RoboDK station: paint_booth.rdk

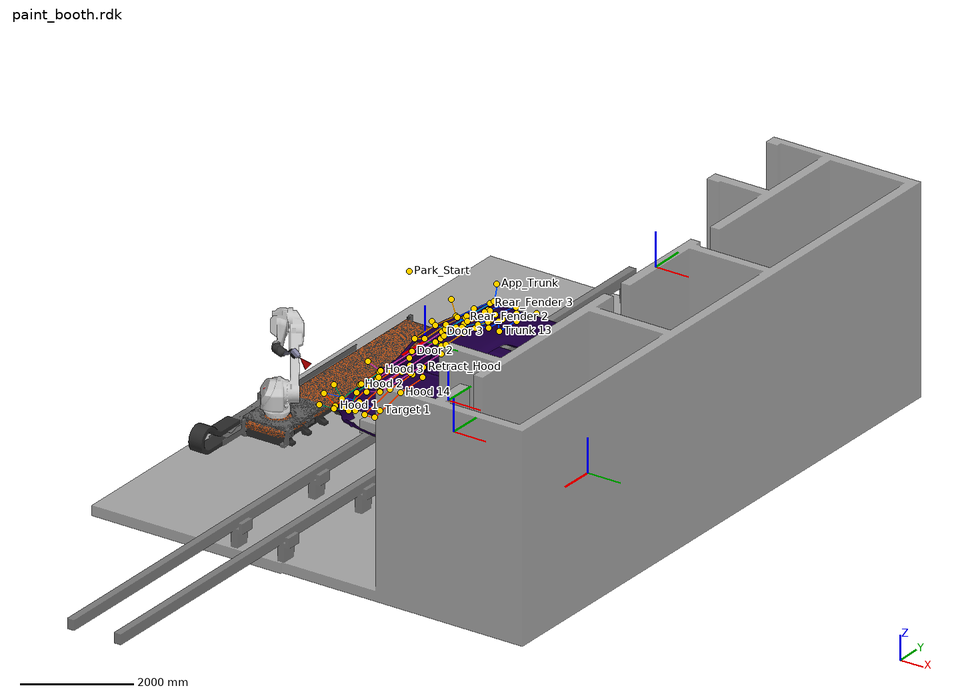
[picture v0: the station drawn from its stored meshes, robots at their saved joint values, targets as dots, program paths as lines]
Station paint booth backup2 (saved by RoboDK 6.1.1). Poses are relative to the parent item; angles as X-Y-Z fixed-axis rotations.
Station parameters (name, value as stored): AttachCamera_Record, 1, Record_Record, 0
  - frame ABB IRBT 7004 Standard 4m Base at (0, 2700, 0) mm, rotated rx 0 ry 0 rz -90 deg
    - robot ABB IRBT 7004 Standard 4m: 1 axes
        modified DH rows (alpha deg, a mm, theta deg, d mm): 0, 0, 0, 0 linear
        base shift (840.5, 4.2, 379.5) mm, rotated rx 0 ry 90 rz 0 deg
        joint limits [0] to [3700]; home [0]; saved at [3700]
      - robot ABB IRB 5500-27: 6 axes, payload 16 kg, reach 2200 mm, repeatability 0.15 mm, weight 600 kg
          modified DH rows (alpha deg, a mm, theta deg, d mm): 0, 0, 0, 436; -90, 0, -90, -5; 0, 1300, 0, 0; -90, 0, -90, 1510.5; 35, 0, 0, 79.169; -70, 0, 180, 79.169
          base shift (0, 0, 0) mm, rotated rx 0 ry 0 rz 90 deg
          joint limits [-104, -65, -70, -719, -719, -720] to [104, 150, 70, 719, 719, 720]; home [0, 0, 0, 0, 0, 0]; saved at [-54.839, -32.896, 27.054, 12.85, -64.516, 53.554]
        - tool Generic Paint Sprayer, TCP at (87.9, 0, 515.6) mm, rotated rx 0 ry 30 rz 0 deg, size 277.6 x 203.2 x 501.7 mm
  - frame booth_frame at (5380, 0, 0) mm, rotated rx 0 ry 0 rz -90 deg
    - folder Paint_Booth
      - object paint booth v1_paint booth v1_Back wall at (0, 0, 0) mm, size 12200 x 2000 x 4000 mm, geometry from paint booth v1_paint booth v1_Back wall.stl
      - object paint booth v1_paint booth v1_entry_part at (0, 0, 0) mm, size 250 x 1150 x 4000 mm, geometry from paint booth v1_paint booth v1_entry_part.stl
      - object paint booth v1_paint booth v1_entry_wall (1) at (0, 0, 0) mm, size 250 x 1150 x 4000 mm, geometry from paint booth v1_paint booth v1_entry_wall (1).stl
      - object paint booth v1_paint booth v1_entry_wall at (0, 0, 0) mm, size 1700 x 439.1 x 4000 mm, geometry from paint booth v1_paint booth v1_entry_wall.stl
      - object paint booth v1_paint booth v1_exit_wall (1) at (0, 0, 0) mm, size 250 x 1150 x 4000 mm, geometry from paint booth v1_paint booth v1_exit_wall (1).stl
      - object paint booth v1_paint booth v1_exit_wall (2) at (0, 0, 0) mm, size 250 x 1150 x 4000 mm, geometry from paint booth v1_paint booth v1_exit_wall (2).stl
      - object paint booth v1_paint booth v1_exit_wall at (0, 0, 0) mm, size 2500 x 439.1 x 4000 mm, geometry from paint booth v1_paint booth v1_exit_wall.stl
      - object paint booth v1_paint booth v1_floor at (0, 0, 0) mm, size 12240.8 x 9200 x 200 mm, geometry from paint booth v1_paint booth v1_floor.stl
      - object paint booth v1_paint booth v1_front_wall at (0, 0, 0) mm, size 8000 x 200 x 4000 mm, geometry from paint booth v1_paint booth v1_front_wall.stl
      - object paint booth v1_paint booth v1_mid_wall (1) at (0, 0, 0) mm, size 4000 x 200 x 4000 mm, geometry from paint booth v1_paint booth v1_mid_wall (1).stl
      - object paint booth v1_paint booth v1_mid_wall (2) at (0, 0, 0) mm, size 950 x 200 x 4000 mm, geometry from paint booth v1_paint booth v1_mid_wall (2).stl
      - object paint booth v1_paint booth v1_mid_wall (3) at (0, 0, 0) mm, size 3400 x 200 x 4000 mm, geometry from paint booth v1_paint booth v1_mid_wall (3).stl
      - object paint booth v1_paint booth v1_mid_wall at (0, 0, 0) mm, size 2150 x 200 x 4000 mm, geometry from paint booth v1_paint booth v1_mid_wall.stl
  - frame conveyor_frame at (2500, 0, 0) mm
    - object Conveyor at (0, 6191.19, 0) mm, rotated rx 0 ry 0 rz -90 deg, size 17200 x 1350 x 600 mm, geometry from Conveyor.stl
    - object cart at (0, 6191.19, 0) mm, size 1500 x 3500 x 250 mm, geometry from cart.stl
    - frame frame_base at (0, 6191.19, 750) mm
    - target Conv_Entry (joint target) at (0, 1691.19, 750) mm; joints [0] of Conveyor
    - target Conv_Paint (joint target) at (0, 1691.19, 750) mm; joints [4500] of Conveyor
    - target Conv_Exit (joint target) at (0, 1691.19, 750) mm; joints [13248.192] of Conveyor
  - frame Conveyor at (2500, 6191.19, 750) mm
    - robot Conveyor: 1 axes
        modified DH rows (alpha deg, a mm, theta deg, d mm): 0, 0, 0, 0 linear
        base shift (0, 0, 0) mm, rotated rx 90 ry 0 rz 0 deg
        joint limits [0] to [15000]; home [0]; saved at [4500]
      - frame car_frame at (0, -1850, -70) mm
        - object car_body at (0, 0, 0) mm, rotated rx 90 ry 0 rz 90 deg, size 4801.1 x 1114.9 x 1961.6 mm, geometry from car_body_optimised.obj
        - target Target 1 (Cartesian target) at (20.58, -2128.6, 648.13) mm, rotated rx 159.32 ry 5.46 rz -156.1 deg; joints [-17.994, 40.195, -43.091, -41.526, -55.736, 93.269, 3700] of ABB IRB 5500-27
        - target Target 2 (Cartesian target) at (-499.07, -2013.93, 637.53) mm, rotated rx 169.55 ry 9.47 rz -156.84 deg; joints [-17.854, 10.002, -1.972, -48.865, -37.872, 74.599, 3700] of ABB IRB 5500-27
        - object car_paint_1 at (-2500, 158.81, -680) mm, size 1941.7 x 1314.7 x 689.4 mm
        - object car_paint_2 at (-2500, 158.81, -680) mm, size 1932.4 x 3061.3 x 1113.1 mm
        - object car_paint_3 at (-2500, 158.81, -680) mm, size 1960.3 x 2051 x 1094.9 mm
        - object car_paint_4 at (-2500, 158.81, -680) mm, size 1961.6 x 1256.6 x 838.3 mm
        - target Hood 1 (Cartesian target) at (-850, -2240, 549.52) mm, rotated rx 170.58 ry 46.52 rz 180 deg; joints [-33.908, -9.39, 33.602, 38.78, -64.314, 10.994, 3700] of ABB IRB 5500-27
        - target Hood 2 (Cartesian target) at (-850, -1495, 668.46) mm, rotated rx 175.62 ry 0.84 rz -135.11 deg; joints [-8.251, -3.639, 8.764, -39.401, -59.237, 68.878, 3513] of ABB IRB 5500-27
        - target Hood 3 (Cartesian target) at (-850, -850, 690.55) mm, rotated rx 179.29 ry 0.3 rz -135 deg; joints [-7.072, -4.967, 9.136, -44.55, -55.783, 68.456, 2868] of ABB IRB 5500-27
        - target Hood 4 (Cartesian target) at (-625, -850, 729.52) mm, rotated rx -176.51 ry 5.77 rz -134.73 deg; joints [-6.745, 1.906, 2.143, -43.43, -50.492, 62.325, 2868] of ABB IRB 5500-27
        - target Hood 5 (Cartesian target) at (-625, -1505, 702.48) mm, rotated rx 179.51 ry 6.71 rz -134.83 deg; joints [-8.01, 3.25, 1.791, -36.982, -54.709, 62.353, 3523] of ABB IRB 5500-27
        - target Hood 6 (Cartesian target) at (-625, -2260, 584.84) mm, rotated rx 153.99 ry 5.37 rz -180 deg; joints [-27.175, 8.933, 2.732, -74.826, -17.731, 103.498, 3700] of ABB IRB 5500-27
        - target Hood 7 (Cartesian target) at (-400, -2280, 595.96) mm, rotated rx 166.53 ry -24.84 rz 109.32 deg; joints [-16.554, 21.687, -16.957, -133.314, -63.434, 218.22, 3700] of ABB IRB 5500-27
        - target Hood 8 (Cartesian target) at (-400, -1515, 725.47) mm, rotated rx 177.2 ry 3.28 rz 134.91 deg; joints [6.733, 12.58, -7.202, -178.41, -50.579, 227.726, 3533] of ABB IRB 5500-27
        - target Hood 9 (Cartesian target) at (-400, -850, 782.15) mm, rotated rx 177.63 ry 2.98 rz 134.92 deg; joints [6.843, 12.694, -9.476, -174.35, -52.852, 224.109, 2868] of ABB IRB 5500-27
        - target Hood 10 (Cartesian target) at (-175, -850, 793.95) mm, rotated rx 179.19 ry 2.16 rz 134.97 deg; joints [6.345, 23.93, -24.263, -167.605, -56.502, 217.205, 2868] of ABB IRB 5500-27
        - target Hood 11 (Cartesian target) at (-175, -1535, 771.67) mm, rotated rx 175.02 ry -3.19 rz 135.2 deg; joints [4.513, 24.031, -24.527, -162.354, -53.815, 216.084, 3553] of ABB IRB 5500-27
        - target Hood 12 (Cartesian target) at (-175, -2320, 594.33) mm, rotated rx 153.88 ry -17.93 rz 140.44 deg; joints [-26.584, 35.128, -33.541, -146.9, -20.302, 192.59, 3400] of ABB IRB 5500-27
        - target Retract_Hood (Cartesian target) at (51.74, -845.07, 996.33) mm, rotated rx -178.53 ry 0.28 rz 150.01 deg; joints [4.772, 37.088, -50.956, -153.474, -51.155, 189.496, 2868] of ABB IRB 5500-27
        - target App_Hood (Cartesian target) at (-1064.75, -2289.09, 753.16) mm, rotated rx 170.58 ry 46.52 rz 180 deg; joints [-42.072, -20.414, 34.025, 25.717, -61.677, 26.626, 3700] of ABB IRB 5500-27
        - target Hood 13 (Cartesian target) at (50, -2320, 604.2) mm, rotated rx 153.39 ry -19.8 rz 153.35 deg; joints [-18.538, 44.698, -49.255, -115.628, -40.633, 174.214, 3700] of ABB IRB 5500-27
        - target Hood 14 (Cartesian target) at (50, -1535, 774.22) mm, rotated rx 175.67 ry -3.9 rz 150.09 deg; joints [2.571, 34.693, -39.712, -165.563, -37, 201.31, 3553] of ABB IRB 5500-27
        - target Hood 15 (Cartesian target) at (50, -850, 796.4) mm, rotated rx -178.53 ry 0.28 rz 150.01 deg; joints [4.294, 34.498, -39.52, -172.584, -37.994, 202.13, 2868] of ABB IRB 5500-27
        - target App_Fender (Cartesian target) at (-974.76, -2108.13, 875.32) mm, rotated rx 153.92 ry -10.06 rz 94.89 deg; joints [-22.913, -9.502, 9.705, -153.801, -59.777, 240.063, 3400] of ABB IRB 5500-27
        - target Fender 1 (Cartesian target) at (-847.37, -2050, 610) mm, rotated rx 153.92 ry -10.06 rz 94.89 deg; joints [-6.967, -7.664, 17.735, -150.991, -72.848, 258.721, 3700] of ABB IRB 5500-27
        - target Fender 2 (Cartesian target) at (-906.3, -1375, 610) mm, rotated rx 112.74 ry -29.02 rz 81.54 deg; joints [-2.631, -20.422, 36.583, -152.192, -69.948, 315.942, 3093] of ABB IRB 5500-27
        - target Fender 3 (Cartesian target) at (-916.58, -800, 610) mm, rotated rx 111.21 ry -14.19 rz 85.06 deg; joints [-0.206, -20.739, 39.32, -164.713, -74.487, 320.113, 2518] of ABB IRB 5500-27
        - target Fender 4 (Cartesian target) at (-964.37, -800, 470) mm, rotated rx 83.95 ry -44.78 rz 95.04 deg; joints [13.122, -20.802, 49.517, -168.289, -57.057, 363.142, 2818] of ABB IRB 5500-27
        - target Fender 5 (Cartesian target) at (-947.24, -1462.5, 470) mm, rotated rx 78.8 ry -44.05 rz 100.71 deg; joints [11.072, -19.709, 50.508, -183.586, -47.435, 370.499, 3480.5] of ABB IRB 5500-27
        - target Fender 6 (Cartesian target) at (-892.02, -2225, 470) mm, rotated rx 90.97 ry -0.07 rz 94.26 deg; joints [-18.235, -10.576, 47.923, -230.993, -54.777, 371.88, 3700] of ABB IRB 5500-27
        - target Retract_Fender (Cartesian target) at (-1191.15, -2247.27, 475.09) mm, rotated rx 90.97 ry -0.07 rz 94.26 deg; joints [-27.587, -27.313, 58.426, -256.591, -35.126, 378.189, 3700] of ABB IRB 5500-27
        - target Fender 8 (Cartesian target) at (-931.33, -765.59, 218.07) mm, rotated rx 72.26 ry -43.35 rz 102.38 deg; joints [11.704, -5.54, 53.432, -204.915, -44.004, 400.952, 2783.594] of ABB IRB 5500-27
        - target Fender 7 (Cartesian target) at (-891.01, -1776.07, 252.43) mm, rotated rx 71.68 ry -38.06 rz 103.98 deg; joints [4.854, -4.611, 52.488, -218.536, -40.98, 403.383, 3700] of ABB IRB 5500-27
        - target App_Door (Cartesian target) at (-1193.57, -760.98, 726.36) mm, rotated rx 118.17 ry 41.33 rz 109.68 deg; joints [-11.246, -41.025, 55.296, -250.139, -53.107, 329.229, 2478] of ABB IRB 5500-27
        - target Door 1 (Cartesian target) at (-913.06, -760, 620) mm, rotated rx 118.17 ry 41.33 rz 109.68 deg; joints [-7.482, -20.017, 48.249, -231.788, -76.441, 333.571, 2478] of ABB IRB 5500-27
        - target Door 2 (Cartesian target) at (-912.63, 190, 620) mm, rotated rx 118.57 ry 41.24 rz 109.9 deg; joints [-7.46, -20.08, 48.148, -232.112, -75.877, 333.185, 1528] of ABB IRB 5500-27
        - target Door 3 (Cartesian target) at (-933.28, 1140, 620) mm, rotated rx 105.5 ry 14.01 rz 95.69 deg; joints [-2.844, -21.627, 47.142, -203.396, -73.018, 334.956, 578] of ABB IRB 5500-27
        - target Door 4 (Cartesian target) at (-963.16, 1140, 480) mm, rotated rx 83.93 ry -44.87 rz 93.9 deg; joints [13.914, -20.65, 48.974, -164.88, -60.023, 363.185, 878] of ABB IRB 5500-27
        - target Door 5 (Cartesian target) at (-965.98, 190, 480) mm, rotated rx 87.35 ry -44.97 rz 91.86 deg; joints [13.842, -21.244, 48.306, -160.437, -62.168, 358.751, 1828] of ABB IRB 5500-27
        - target Door 6 (Cartesian target) at (-965.55, -760, 480) mm, rotated rx 85.39 ry -44.87 rz 93.85 deg; joints [13.359, -21.255, 48.945, -164.795, -59.171, 360.752, 2778] of ABB IRB 5500-27
        - target Door 7 (Cartesian target) at (-952.18, -760, 340) mm, rotated rx 82.3 ry -29.74 rz 94.11 deg; joints [15.675, -11.351, 52.057, -173.644, -71.818, 377.792, 2778] of ABB IRB 5500-27
        - target Door 8 (Cartesian target) at (-952.1, 190, 340) mm, rotated rx 81.98 ry -29.77 rz 93.93 deg; joints [15.886, -11.116, 52.001, -173.048, -72.449, 378.36, 1828] of ABB IRB 5500-27
        - target Door 9 (Cartesian target) at (-950.94, 1140, 340) mm, rotated rx 83.74 ry -29.64 rz 95.3 deg; joints [14.421, -12.419, 52.327, -177.488, -68.067, 375.266, 878] of ABB IRB 5500-27
        - target Door 10 (Cartesian target) at (-934.75, 1120, 200) mm, rotated rx 85.21 ry 3.16 rz 123.35 deg; joints [-7.502, 0.911, 55.483, -244.469, -73.616, 400.866, 898] of ABB IRB 5500-27
        - target Door 11 (Cartesian target) at (-927.07, 180, 200) mm, rotated rx 71.8 ry -43.53 rz 102.75 deg; joints [11.512, -4.316, 53.386, -207.144, -43.231, 403.245, 1838] of ABB IRB 5500-27
        - target Door 12 (Cartesian target) at (-927.11, -760, 200) mm, rotated rx 71.28 ry -43.44 rz 103.11 deg; joints [11.489, -4.115, 53.426, -207.745, -43.268, 404.073, 2778] of ABB IRB 5500-27
        - target Retract_Door (Cartesian target) at (-1218.85, -759.98, 130.1) mm, rotated rx 71.28 ry -43.44 rz 103.11 deg; joints [16.969, -15.398, 66.274, -198.158, -49.917, 404.175, 2778] of ABB IRB 5500-27
        - target App_Rear_Fender (Cartesian target) at (-1226.32, 1241.64, 697.15) mm, rotated rx -104.9 ry 0.41 rz -88.46 deg; joints [24.298, -37.224, 47.754, -398.951, -32.669, 337.437, 1368] of ABB IRB 5500-27
        - target Rear_Fender 1 (Cartesian target) at (-936.54, 1250, 620) mm, rotated rx -104.9 ry 0.41 rz -88.46 deg; joints [17.106, -19.16, 39.645, -373.877, -49.209, 317.907, 1368] of ABB IRB 5500-27
        - target Rear_Fender 2 (Cartesian target) at (-930.4, 1850, 620) mm, rotated rx -110.85 ry -0.76 rz -91.99 deg; joints [2.229, -22.32, 39.28, -367.971, -67.352, 327.123, 468] of ABB IRB 5500-27
        - target Rear_Fender 3 (Cartesian target) at (-899.38, 2550, 620) mm, rotated rx -131.31 ry 33.88 rz -121.93 deg; joints [20.837, -18.952, 39.054, -347.896, -25.853, 323.447, 0] of ABB IRB 5500-27
        - target Rear_Fender 4 (Cartesian target) at (-940.1, 2550, 480) mm, rotated rx -86.44 ry -14.81 rz -93.66 deg; joints [17.494, -14.594, 46.728, -380.009, -36.647, 287.127, 0] of ABB IRB 5500-27
        - target Rear_Fender 5 (Cartesian target) at (-958.49, 1850, 480) mm, rotated rx -85.17 ry -29.81 rz -93.81 deg; joints [-13.408, -18.273, 46.663, -377.953, -71.976, 283.944, 168] of ABB IRB 5500-27
        - target Rear_Fender 6 (Cartesian target) at (-963.3, 1250, 480) mm, rotated rx -85.81 ry -44.94 rz -92.57 deg; joints [-10.68, -20.846, 45.763, -404.205, -59.45, 290.619, 768] of ABB IRB 5500-27
        - target Rear_Fender 7 (Cartesian target) at (-960.41, 1840, 300) mm, rotated rx 70.16 ry -59.4 rz 101.96 deg; joints [9.883, -14.191, 50.692, -282.824, 27.785, 438.94, 178] of ABB IRB 5500-27
        - target Rear_Fender 8 (Cartesian target) at (-926.34, 2140, 300) mm, rotated rx 59.88 ry -57.09 rz 113.2 deg; joints [15.432, -9.247, 49.626, -292.317, 26.354, 453.547, 0] of ABB IRB 5500-27
        - target Rear_Fender 9 (Cartesian target) at (-880.15, 2540, 300) mm, rotated rx 13.56 ry -52.4 rz 131.86 deg; joints [39.466, 17.311, 30.479, -344.467, 73.043, 520.699, 0] of ABB IRB 5500-27
        - target Retract_Rear_Fender (Cartesian target) at (-1214.63, 2153.98, 218.19) mm, rotated rx 59.88 ry -57.09 rz 113.2 deg; joints [23.086, -20.703, 61.466, -305.303, 38.947, 463.966, 0] of ABB IRB 5500-27
        - target App_Roof (Cartesian target) at (-25.83, 1302.61, 1216.86) mm, rotated rx -162.4 ry 4.89 rz 165.72 deg; joints [7.333, 34.052, -54.57, -280.864, 45.422, 591.934, 778] of ABB IRB 5500-27
        - target Roof 1 (Cartesian target) at (-700, -40, 1021.33) mm, rotated rx -137.85 ry 38.85 rz -115.76 deg; joints [-11.875, -13.9, 23.29, -152.293, 73.605, 433.224, 2058] of ABB IRB 5500-27
        - target Roof 2 (Cartesian target) at (-700, 600, 1031.86) mm, rotated rx -134.41 ry 21.13 rz -111.88 deg; joints [-10.086, -13.722, 18.402, -167.792, 67.736, 438.526, 1418] of ABB IRB 5500-27
        - target Roof 3 (Cartesian target) at (-700, 1240, 956.24) mm, rotated rx -144.33 ry 3.95 rz -123.41 deg; joints [-2.958, -10.964, 12.354, -168.948, 40.63, 457.779, 778] of ABB IRB 5500-27
        - target Roof 4 (Cartesian target) at (-475, 1240, 1022.67) mm, rotated rx -163.75 ry -7.87 rz -151.31 deg; joints [1.04, 8.492, -14.517, -201.236, 31.187, 517.343, 778] of ABB IRB 5500-27
        - target Roof 5 (Cartesian target) at (-475, 600, 1103.28) mm, rotated rx -177.98 ry 1.17 rz -150 deg; joints [-4.572, 8.746, -17.039, -191.609, 39.597, 518.656, 1418] of ABB IRB 5500-27
        - target Roof 6 (Cartesian target) at (-475, -40, 1082.57) mm, rotated rx 166.05 ry 11.35 rz -150.93 deg; joints [-10.13, 8.919, -13.503, -173.375, 44.185, 514.846, 2058] of ABB IRB 5500-27
        - target Roof 7 (Cartesian target) at (-250, -40, 1090.04) mm, rotated rx 161.81 ry -3.66 rz 165.76 deg; joints [-3.903, 18.259, -27.873, -207.606, 15.657, 578.393, 2058] of ABB IRB 5500-27
        - target Roof 8 (Cartesian target) at (-250, 600, 1108.78) mm, rotated rx -178.57 ry 1.25 rz 165 deg; joints [1.727, 18.57, -29.817, -240.694, 22.465, 586.685, 1418] of ABB IRB 5500-27
        - target Roof 9 (Cartesian target) at (-250, 1240, 1025.03) mm, rotated rx -162.62 ry 5.04 rz 165.7 deg; joints [6.33, 18.4, -25.159, -256.892, 18.962, 589.513, 778] of ABB IRB 5500-27
        - target Roof 10 (Cartesian target) at (-25, 1240, 1026.91) mm, rotated rx -162.4 ry 4.89 rz 165.72 deg; joints [5.697, 30.2, -41.291, -263.996, 27.262, 589.828, 778] of ABB IRB 5500-27
        - target Roof 11 (Cartesian target) at (-25, 600, 1111.34) mm, rotated rx -178.33 ry 0.61 rz 165.01 deg; joints [1.451, 31.512, -48.022, -254.939, 35.89, 591.02, 1418] of ABB IRB 5500-27
        - target Roof 12 (Cartesian target) at (-25, -40, 1092.94) mm, rotated rx 162.68 ry -4.28 rz 165.69 deg; joints [-3.688, 31.077, -45.986, -232.063, 33.174, 590.485, 2058] of ABB IRB 5500-27
        - target Retract_Roof (Cartesian target) at (-855.26, 1322.31, 1199.39) mm, rotated rx -144.33 ry 3.95 rz -123.41 deg; joints [0.151, -16.974, 8.301, -182.475, 44.016, 473.293, 778] of ABB IRB 5500-27
        - target App_Trunk (Cartesian target) at (-871.24, 2723.68, 933.63) mm, rotated rx -159.78 ry 4.33 rz 180 deg; joints [34.013, 0.121, -2.145, -300.577, 42.076, 618.392, 0] of ABB IRB 5500-27
        - target Trunk 1 (Cartesian target) at (-850, 1480, 788.68) mm, rotated rx 176.99 ry 6.8 rz 134.66 deg; joints [8.818, -8.186, 9.746, -321.801, 55.89, 657.36, 538] of ABB IRB 5500-27
        - target Trunk 2 (Cartesian target) at (-850, 2000, 748.95) mm, rotated rx -176.67 ry 4.21 rz 135.09 deg; joints [9.552, -5.157, 7.83, -325.039, 61.252, 652.551, 18] of ABB IRB 5500-27
        - target Trunk 3 (Cartesian target) at (-850, 2620, 652.92) mm, rotated rx -159.78 ry 4.33 rz 180 deg; joints [30.207, -0.765, 9.349, -286.741, 23.622, 619.899, 0] of ABB IRB 5500-27
        - target Trunk 4 (Cartesian target) at (-625, 2640, 651.31) mm, rotated rx -160.39 ry 0.99 rz -180 deg; joints [26.359, 9.187, -1.352, -266.924, 15.228, 605.429, 0] of ABB IRB 5500-27
        - target Trunk 5 (Cartesian target) at (-625, 2010, 751.36) mm, rotated rx -176.73 ry 4.49 rz 135.09 deg; joints [8.299, 4.538, -1.818, -323.121, 59.025, 651.92, 8] of ABB IRB 5500-27
        - target Trunk 6 (Cartesian target) at (-625, 1480, 769.14) mm, rotated rx 178.96 ry -1.18 rz 135.01 deg; joints [5.561, 4.409, -3.241, -310.888, 55.555, 647.783, 538] of ABB IRB 5500-27
        - target Trunk 7 (Cartesian target) at (-400, 1480, 768.9) mm, rotated rx 178.96 ry -1.12 rz 135.01 deg; joints [4.907, 14.354, -14.487, -310.139, 55.784, 646.085, 538] of ABB IRB 5500-27
        - target Trunk 8 (Cartesian target) at (-400, 2010, 754.63) mm, rotated rx -176.58 ry 4.39 rz 135.1 deg; joints [7.289, 14.473, -13.215, -321.436, 58.548, 649.531, 8] of ABB IRB 5500-27
        - target Trunk 9 (Cartesian target) at (-400, 2640, 654.71) mm, rotated rx -162.66 ry 10.33 rz 151.49 deg; joints [27.495, 22.985, -18.315, -343.977, 71.386, 648.375, 0] of ABB IRB 5500-27
        - target Trunk 10 (Cartesian target) at (-175, 2340, 717.22) mm, rotated rx -174.44 ry 6.26 rz 135.27 deg; joints [15.939, 28.451, -29.809, -338.469, 74.927, 651.2, 0] of ABB IRB 5500-27
        - target Trunk 11 (Cartesian target) at (-175, 1910, 766.78) mm, rotated rx -176.59 ry 4.27 rz 135.1 deg; joints [6.472, 24.893, -26.972, -320.217, 59.841, 645.622, 108] of ABB IRB 5500-27
        - target Trunk 12 (Cartesian target) at (-175, 1480, 768.85) mm, rotated rx 178.96 ry -1.04 rz 135.01 deg; joints [4.405, 24.857, -27.881, -310.287, 57.894, 643.265, 538] of ABB IRB 5500-27
        - target Retract_Trunk (Cartesian target) at (50.01, 1474.88, 968.79) mm, rotated rx 178.96 ry -1.04 rz 135.01 deg; joints [3.942, 39.672, -56.806, -316.42, 72.72, 631.534, 538] of ABB IRB 5500-27
        - target Trunk 13 (Cartesian target) at (50, 1480, 768.86) mm, rotated rx 178.96 ry -1.04 rz 135.01 deg; joints [4.004, 36.972, -45.172, -311.787, 62.792, 638.73, 538] of ABB IRB 5500-27
        - target Trunk 14 (Cartesian target) at (50, 2010, 758.1) mm, rotated rx -175.81 ry 3.84 rz 135.15 deg; joints [5.895, 37.28, -44.398, -320.475, 63.909, 639.675, 8] of ABB IRB 5500-27
        - target Trunk 15 (Cartesian target) at (50, 2640, 656.35) mm, rotated rx -161.94 ry 10.12 rz 151.62 deg; joints [22.605, 44.732, -49.956, -335.396, 68.161, 635.183, 0] of ABB IRB 5500-27
        - target Park_Start (joint target) at (-1755.26, 1322.31, 1499.39) mm, rotated rx -144.33 ry 3.95 rz -123.41 deg; joints [-54.839, -32.896, 27.054, 12.85, -64.516, 53.554, 3700] of ABB IRB 5500-27
        - target Park_End (joint target) at (-1755.26, 1322.31, 1499.39) mm, rotated rx -144.33 ry 3.95 rz -123.41 deg; joints [53.695, -43.794, 10.536, -128.115, -49.304, 481.516, 1078] of ABB IRB 5500-27
  - program Prog2 (10 instructions, listed below)
  - program Paint_Hood (31 instructions, listed below)
  - program Paint_Fender (19 instructions, listed below)
  - program Paint_Door (26 instructions, listed below)
  - program Paint_Roof (26 instructions, listed below)
  - program Paint_Rear_Fender (21 instructions, listed below)
  - program Paint_Trunk (31 instructions, listed below)
  - program Main_Paint (7 instructions, listed below)
  - Python program SprayOn (listed below)
  - program Robot_Park_Start (2 instructions, listed below)
  - program Robot_Park_End (2 instructions, listed below)
  - program Conveyor_Reset (2 instructions, listed below)
  - program Conveyor_In (2 instructions, listed below)
  - program Conveyor_Out (2 instructions, listed below)
  - program Cell_Cycle (6 instructions, listed below)
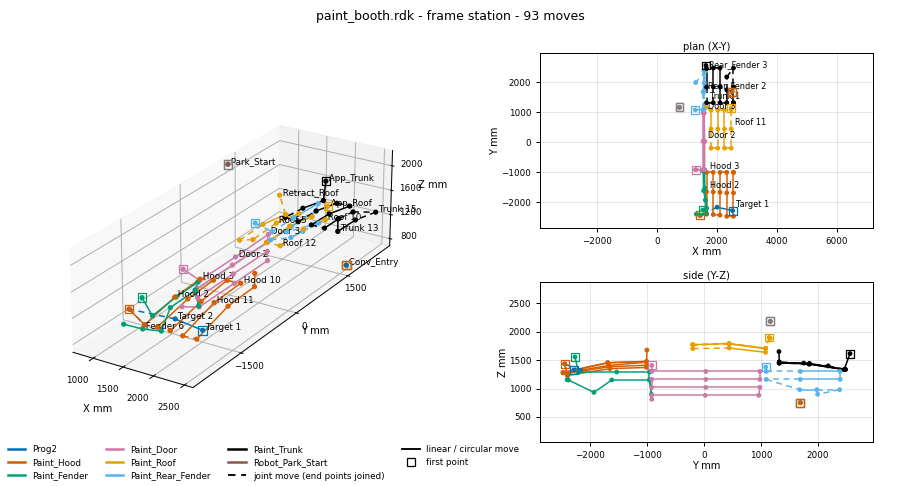
[picture p0: tool path of paint_booth.rdk in frame station, 93 of 93 moves have a stored position in this frame; points joined in program order, loops and branches not executed]

--- program Prog2 (robot ABB IRB 5500-27) ---
  Set Ref.: car_frame
  Set Tool: Generic Paint Sprayer
  Call SprayOn(-1)
  MoveJ (Target 1)
  Set speed (500.0 mm/s)
  Call SprayOn(1)
  MoveL (Target 2)
  Call SprayOn(0)
  MoveJ (App_Hood)
  MoveJ (Hood 1)

--- program Paint_Hood (robot ABB IRB 5500-27) ---
  Set Ref.: car_frame
  Set Tool: Generic Paint Sprayer
  Set speed (1000.0 mm/s)
  MoveJ (App_Hood)
  Set speed (500.0 mm/s)
  MoveL (Hood 1)
  Call SprayOn(1)
  MoveL (Hood 2)
  MoveL (Hood 3)
  Call SprayOn(0)
  MoveJ (Hood 4)
  Call SprayOn(1)
  MoveL (Hood 5)
  MoveL (Hood 6)
  Call SprayOn(0)
  MoveJ (Hood 7)
  Call SprayOn(1)
  MoveL (Hood 8)
  MoveL (Hood 9)
  Call SprayOn(0)
  MoveJ (Hood 10)
  Call SprayOn(1)
  MoveL (Hood 11)
  MoveL (Hood 12)
  Call SprayOn(0)
  MoveJ (Hood 13)
  Call SprayOn(1)
  MoveL (Hood 14)
  MoveL (Hood 15)
  Call SprayOn(0)
  MoveL (Retract_Hood)

--- program Paint_Fender (robot ABB IRB 5500-27) ---
  Set Ref.: car_frame
  Set Tool: Generic Paint Sprayer
  Set speed (1000.0 mm/s)
  MoveJ (App_Fender)
  Set speed (500.0 mm/s)
  MoveL (Fender 1)
  Call SprayOn(1)
  MoveL (Fender 2)
  MoveL (Fender 3)
  Call SprayOn(0)
  MoveJ (Fender 4)
  Call SprayOn(1)
  MoveL (Fender 8)
  MoveL (Fender 4)
  MoveL (Fender 5)
  MoveL (Fender 7)
  MoveL (Fender 6)
  Call SprayOn(0)
  MoveL (Retract_Fender)

--- program Paint_Door (robot ABB IRB 5500-27) ---
  Set Ref.: car_frame
  Set Tool: Generic Paint Sprayer
  Set speed (1000.0 mm/s)
  MoveJ (App_Door)
  Set speed (500.0 mm/s)
  MoveL (Door 1)
  Call SprayOn(1)
  MoveL (Door 2)
  MoveL (Door 3)
  Call SprayOn(0)
  MoveJ (Door 4)
  Call SprayOn(1)
  MoveL (Door 5)
  MoveL (Door 6)
  Call SprayOn(0)
  MoveJ (Door 7)
  Call SprayOn(1)
  MoveL (Door 8)
  MoveL (Door 9)
  Call SprayOn(0)
  MoveJ (Door 10)
  Call SprayOn(1)
  MoveL (Door 11)
  MoveL (Door 12)
  Call SprayOn(0)
  MoveL (Retract_Door)

--- program Paint_Roof (robot ABB IRB 5500-27) ---
  Set Ref.: car_frame
  Set Tool: Generic Paint Sprayer
  Set speed (1000.0 mm/s)
  MoveJ (App_Roof)
  Set speed (500.0 mm/s)
  MoveJ (Roof 10)
  Call SprayOn(1)
  MoveJ (Roof 11)
  MoveJ (Roof 12)
  Call SprayOn(0)
  MoveJ (Roof 7)
  Call SprayOn(1)
  MoveL (Roof 8)
  MoveL (Roof 9)
  Call SprayOn(0)
  MoveJ (Roof 4)
  Call SprayOn(1)
  MoveL (Roof 5)
  MoveJ (Roof 6)
  Call SprayOn(0)
  MoveJ (Roof 1)
  Call SprayOn(1)
  MoveJ (Roof 2)
  MoveL (Roof 3)
  Call SprayOn(0)
  MoveJ (Retract_Roof)

--- program Paint_Rear_Fender (robot ABB IRB 5500-27) ---
  Set Ref.: car_frame
  Set Tool: Generic Paint Sprayer
  Set speed (1000.0 mm/s)
  MoveJ (App_Rear_Fender)
  Set speed (500.0 mm/s)
  MoveJ (Rear_Fender 1)
  Call SprayOn(1)
  MoveJ (Rear_Fender 2)
  MoveL (Rear_Fender 3)
  Call SprayOn(0)
  MoveJ (Rear_Fender 4)
  Call SprayOn(1)
  MoveL (Rear_Fender 5)
  MoveJ (Rear_Fender 6)
  Call SprayOn(0)
  MoveJ (Rear_Fender 7)
  Call SprayOn(1)
  MoveL (Rear_Fender 8)
  MoveJ (Rear_Fender 9)
  Call SprayOn(0)
  MoveJ (Retract_Rear_Fender)

--- program Paint_Trunk (robot ABB IRB 5500-27) ---
  Set Ref.: car_frame
  Set Tool: Generic Paint Sprayer
  Set speed (1000.0 mm/s)
  MoveJ (App_Trunk)
  Set speed (500.0 mm/s)
  MoveL (Trunk 3)
  Call SprayOn(1)
  MoveL (Trunk 2)
  MoveJ (Trunk 1)
  Call SprayOn(0)
  MoveJ (Trunk 6)
  Call SprayOn(1)
  MoveJ (Trunk 5)
  MoveL (Trunk 4)
  Call SprayOn(0)
  MoveJ (Trunk 9)
  Call SprayOn(1)
  MoveL (Trunk 8)
  MoveL (Trunk 7)
  Call SprayOn(0)
  MoveJ (Trunk 12)
  Call SprayOn(1)
  MoveL (Trunk 11)
  MoveJ (Trunk 10)
  Call SprayOn(0)
  MoveJ (Trunk 15)
  Call SprayOn(1)
  MoveJ (Trunk 14)
  MoveL (Trunk 13)
  Call SprayOn(0)
  MoveL (Retract_Trunk)

--- program Main_Paint (robot ABB IRB 5500-27) ---
  Call SprayOn(-1)
  Call Paint_Hood
  Call Paint_Fender
  Call Paint_Door
  Call Paint_Rear_Fender
  Call Paint_Trunk
  Call Paint_Roof

--- Python program SprayOn ---
# This macro allows simulating a spray gun for painting or to simulate the trace of inspaction
#
# You can call SprayOn(1) to simulate turning the Spray gun ON or SprayOn(0) to stop simulating the gun
# Calling SprayOn(-1) clears all displayed data
# The macro will output spray gun statistics
#
# --------------------------------------------------------------
# This script shows how to create "spray" object in RoboDK that allows simulating particle deposition by using:
# RDK.Spray_Add(tool, object, options_command, volume, geometry)
#    tool: tool item (TCP) to use
#    object: object to project the particles
#    options_command (optional): string to specify options.
#    volume (optional): Matrix of parameters defining the volume of the spray gun
#    geometry (optional): Matrix of vertices defining the triangles.
#
# More information here:
# https://robodk.com/doc/en/PythonAPI/robodk.html#robodk.robolink.Robolink.Spray_Add
# https://robodk.com/doc/en/RoboDK-API.html
#
# The scripts ArcStart, ArcEnd and WeldOn and SpindleOn behave in a similar way, the only difference is the default behavior
# This behavior simmulates Fanuc Arc Welding and triggers appropriate output when using the customized post processor.
# Select ESC to clear the trace manually.
#
# Example scripts that use Spray_Add:
#     SpindleOn / SpindleOff    -> Turn trace On/Off
#     ArcOn / ArcOff            -> Turn trace On/Off
#     SprayOn / SprayOff        -> Simulate a spray given a workspace volume (for painting)
#     WeldOn / WeldOff          -> Support for multiple weld guns

#------------------------------------------------------------------

# Use a specific tool as a spray gun
Tool_Name = 'Generic Paint Sprayer'
#Tool_Name = 'Tool 2'

# Objects to project particles on. The car is split into lengthwise sections
# (car_paint_1..N) because RoboDK's spray projection stopped registering hits
# on a single object spanning the whole 4.8 m car; ~1.2 m sections work.
Object_Prefix = 'car_paint_'
Object_Count = 4

# Process parameters (TCP sits at the standoff point, STANDOFF mm in front of the nozzle)
STANDOFF = 250       # mm, nozzle to painted surface
SPRAY_WIDTH = 300    # mm, spray pattern diameter on the surface
NOZZLE_RADIUS = 15   # mm, cone radius at the nozzle
FAR_OFFSET = 50      # mm, cone extends this far past the surface so particles always hit it

# Define the default action (0 to deactivate, +1 to activate, -1 to clear any spray gun simulation)
# Setting it to None will display a message
ACTION = None

from robodk.robolink import *  # API to communicate with RoboDK
from robodk.robomath import *  # basic matrix operations
from robodk.robodialogs import *

RDK = Robolink()

# quit if we are not in simulation mode
if RDK.RunMode() != RUNMODE_SIMULATE:
    quit()

# Get any previously added spray gun simulations and display statistics (spray on the part vs spray falling out of the part)
info, data = RDK.Spray_GetStats()
if data.size(1) > 0:
    print("Spray gun statistics:")
    print(info)
    print(data.tr())
    # # Diplay statistics
    # RDK.ShowMessage("Material used: %.1f%%<br>Material waisted: %.1f%%<br>Total particles: %.1f" % (data[1,0],data[2,0],data[3,0]), True)
    # # Clear previous spray
    # RDK.Spray_Clear()

# Check if we are running this program inside another program and passing arguments
import sys
if len(sys.argv) > 1:
    ACTION = int(sys.argv[1])

# If the default ACTION is None, display a message to activate/deactivate the spray gun
if ACTION is None:
    print('Note: This macro can be called as Spray(1) or SprayOn(0)')
    entry = mbox('Turn gun ON or OFF', ('On', '1'), ('Off', '0'))
    if not entry:
        quit()
    ACTION = int(entry)

if ACTION == 0:
    # Turn the gun off
    RDK.Spray_SetState(SPRAY_OFF)

elif ACTION < 0:
    # Clear all spray simulations (same as pressing ESC key)
    RDK.Spray_Clear()

elif ACTION > 0 and data.size(1) > 0:
    # The guns already exist (created by an earlier SprayOn(1) in this run):
    # just switch them back on. Adding new ones every pass stacks dozens of
    # simulated guns and stalls the simulation.
    RDK.Spray_SetState(SPRAY_ON)

elif ACTION > 0:
    # First SprayOn(1) after a clear: create the spray gun objects in RoboDK
    # by using RDK.Spray_Add(tool, object, options_command, volume, geometry)
    # tool: tool item (TCP) to use
    # object: object to project the particles
    # options_command (optional): string to specify options. Example:
    #     STEP=AxB: Defines the grid to be projected 1x1 means only one line of particle projection (for example, for welding)
    #     PARTICLE: Defines the shape and size of particle (sphere or particle), unless a specific geometry is provided:
    #       a- SPHERE(radius, facets)
    #       b- SPHERE(radius, facets, scalex, scaley, scalez)
    #       b- CUBE(sizex, sizey, sizez)
    #     RAND=factor: Defines a random factor factor 0 means that the particles are not deposited randomly
    #     ELLYPSE: defines the volume as an ellypse (default)
    #     RECTANGLE: defines the volume as a rectangle
    #     PROJECT: project the particles to the surface (default) (for welding, painting or scanning)
    #     NO_PROJECT: does not project the particles to the surface (for example, for 3D printing)
    #
    # volume (optional): Matrix of parameters defining the volume of the spray gun
    # geometry (optional): Matrix of vertices defining the triangles.

    tool = 0  # auto detect active tool
    obj = 0  # auto detect object in active reference frame
    if Tool_Name is not None:
        tool = RDK.Item(Tool_Name, ITEM_TYPE_TOOL)

    objects = [RDK.Item(Object_Prefix + str(i), ITEM_TYPE_OBJECT) for i in range(1, Object_Count + 1)]
    # We can specify a given tool object and/or object
    #robot = RDK.Item("ABB IRB 2600-12/1.85", ITEM_TYPE_ROBOT)
    #tools = robot.Childs()
    #if len(tools) > 0:
    #    tool = tools[0]
    #obj = RDK.Item('object', ITEM_TYPE_OBJECT)

    options_command = "ELLYPSE PROJECT PARTICLE=SPHERE(10,8,1,1,0.1) STEP=12x12 RAND=8"  # 12x12 grid: light enough for a GTX 1650
    #options_command = "PARTICLE=CUBE(10,10,2) STEP=8x8"
    #options_command = "PARTICLE=SPHERE(4,8) STEP=8x8"
    #options_command = "PARTICLE=SPHERE(4,8,1,1,0.1) STEP=8x8 RAND=3"

    # Example commands for welding:
    # options_command = "PROJECT PARTICLE=SPHERE(4,8)"
    # options_command = PARTICLE=SPHERE(4,8) STEP=1x0

    # define the ellypse volume as p0, pA, pB, colorRGBA (close and far), in mm
    # coordinates must be provided with respect to the TCP
    # Close ellipse at the nozzle, STANDOFF behind the TCP
    close_p0 = [0, 0, -STANDOFF]  # xyz in mm: Center of the conical ellypse (side 1)
    close_pA = [NOZZLE_RADIUS, 0, -STANDOFF]  # xyz in mm: First vertex of the conical ellypse (side 1)
    close_pB = [0, NOZZLE_RADIUS, -STANDOFF]  # xyz in mm: Second vertex of the conical ellypse (side 1)
    close_color = [1, 0, 0, 1]  # RGBA (0-1)

    # Far ellipse FAR_OFFSET past the surface. Similar triangles from the nozzle:
    # radius = (SPRAY_WIDTH/2) * (STANDOFF + FAR_OFFSET) / STANDOFF  -> 150 * 300/250 = 180 mm
    far_radius = (SPRAY_WIDTH / 2) * (STANDOFF + FAR_OFFSET) / STANDOFF
    far_p0 = [0, 0, FAR_OFFSET]  # xyz in mm: Center of the conical ellypse (side 2)
    far_pA = [far_radius, 0, FAR_OFFSET]  # xyz in mm: First vertex of the conical ellypse (side 2)
    far_pB = [0, far_radius, FAR_OFFSET]  # xyz in mm: Second vertex of the conical ellypse (side 2)
    far_color = [0, 0, 1, 0.2]  # RGBA (0-1)

    close_param = close_p0 + close_pA + close_pB + close_color
    far_param = far_p0 + far_pA + far_pB + far_color
    volume = Mat([close_param, far_param]).tr()
    # One simulated gun per car section; they all share the same tool and cone
    for obj in objects:
        RDK.Spray_Add(tool, obj, options_command, volume)
    RDK.Spray_SetState(SPRAY_ON)

    # Another example with a varying rectancular shape
    # define the rectangular volume as p0, pA, pB, colorRGBA (close and far)
    # close_param = [-90,-117,  0,  90,-117,0,   -90,117,  0,       0.2,0.2,1,.1]
    # far_param   = [-175,-190,200, 175,-190,200,   -175,190,200,   0.5,0,0,.9]
    # volume = Mat([close_param, far_param])
    # RDK.Spray_Add(tool, obj, "RECTANGLE PARTICLE=SPHERE(2,5) STEP=15x15 RAND=3", volume.tr())
    # RDK.Spray_SetState(SPRAY_ON)

    # Optional: define geometry as a list of triangles with normals (instead of a scaled cube or a sphere)
    # geom = Mat([[0,0,0,   0,0,1], [5,0,0,   0,0,1], [0,5,0,   0,0,1]])
    # RDK.Spray_Add(tool, obj, "STEP=8x8 RANDX=3", volume.tr(), geom.tr())
    # RDK.Spray_SetState(SPRAY_ON)

--- program Robot_Park_Start (robot ABB IRB 5500-27) ---
  Set speed (1000.0 mm/s)
  MoveJ (Park_Start)

--- program Robot_Park_End (robot ABB IRB 5500-27) ---
  Set speed (1000.0 mm/s)
  MoveJ (Park_End)

--- program Conveyor_Reset (robot Conveyor) ---
  Set speed (3000.0 mm/s)
  MoveJ (Conv_Entry)

--- program Conveyor_In (robot Conveyor) ---
  Set speed (300.0 mm/s)
  MoveJ (Conv_Paint)

--- program Conveyor_Out (robot Conveyor) ---
  Set speed (300.0 mm/s)
  MoveJ (Conv_Exit)

--- program Cell_Cycle (robot ABB IRB 5500-27) ---
  Call Robot_Park_Start
  Call Conveyor_Reset
  Call Conveyor_In
  Call Main_Paint
  Call Robot_Park_End
  Call Conveyor_Out
